(* IEC 61131-3 sources: BODAS-RC27-18_40/st/bodas_rc18_12_27_18_40/plc_logic/application/easyconfig_import/bds_out_ec, 7 files *)

(* ---- bds_out_aov_signal_te-bds_out_aov_signal_te.st ---- *)
(* --- Interface --- *)
{attribute 'qualified_only' := ''}
{attribute 'strict' := ''}
TYPE bds_out_aov_signal_te :
(
	OUT_AOV_START_SIGNALS := 16#300,
	OUT_AOV_START := 16#2FF,
	K25,
	A12,
	K62,
	OUT_AOV_NUM_SIGNALS,
	OUT_AOV_PVG_NUM_SIGNALS := K62
) UINT;
END_TYPE

(* ---- bds_out_do_signal_te-bds_out_do_signal_te.st ---- *)
(* --- Interface --- *)
{attribute 'qualified_only' := ''}
{attribute 'strict' := ''}
TYPE bds_out_do_signal_te :
(
	OUT_DO_START_SIGNALS := 16#100,
	OUT_DO_START := 16#FF,
	K13,
	A04,
	A10,
	A56,
	A11,
	A55,
	A01,
	A06,
	A16,
	A58,
	A49,
	A50,
	K84,
	K85,
	K86,
	K87,
	OUT_DO_NUM_SIGNALS,
	OUT_DO_FSC_NUM_SIGNALS := K84
) UINT;
END_TYPE

(* ---- bds_out_po_signal_te-bds_out_po_signal_te.st ---- *)
(* --- Interface --- *)
{attribute 'qualified_only' := ''}
{attribute 'strict' := ''}
TYPE bds_out_po_signal_te :
(
	OUT_PO_START_SIGNALS := 16#200,
	OUT_PO_START := 16#1FF,
	K07,
	K09,
	K73,
	K08,
	K29,
	K17,
	A32,
	A47,
	A31,
	A48,
	A46,
	A33,
	A34,
	A51,
	A35,
	A53,
	A52,
	A54,
	K16,
	K14,
	K15,
	A19,
	A05,
	A20,
	A09,
	A02,
	A17,
	K51,
	K12,
	A03,
	A18,
	A08,
	A07,
	K80,
	K81,
	K82,
	K83,
	OUT_PO_NUM_SIGNALS,
	OUT_PO_FSC_NUM_SIGNALS := K80,
	OUT_PO_FSC_HS_NUM_SIGNALS := K16
) UINT;
END_TYPE

(* ---- bds_outclcu_signal_te-bds_outClcU_signal_te.st ---- *)
(* --- Interface --- *)
{attribute 'qualified_only' := ''}
{attribute 'strict' := ''}
TYPE bds_outClcU_signal_te :
(
	bds_outClcU_K25_E := 0,
	bds_outClcU_A12_E,
	bds_outClcU_K62_E,
	bds_outClcU_numSignal_E
) USINT;
END_TYPE

(* ---- bds_outdig_signal_te-bds_outDig_signal_te.st ---- *)
(* --- Interface --- *)
{attribute 'external_name' := 'cmp_rts_bds_outDig_signal_te'}
TYPE bds_outDig_signal_te :
(
	bds_outDig_K13_E := 0,
	bds_outDig_A04_E,
	bds_outDig_A10_E,
	bds_outDig_A56_E,
	bds_outDig_A11_E,
	bds_outDig_A55_E,
	bds_outDig_A01_E,
	bds_outDig_A06_E,
	bds_outDig_A16_E,
	bds_outDig_A58_E,
	bds_outDig_A49_E,
	bds_outDig_A50_E,
	bds_outDig_K84_E,
	bds_outDig_K85_E,
	bds_outDig_K86_E,
	bds_outDig_K87_E,
	bds_outDig_K07_E,
	bds_outDig_K09_E,
	bds_outDig_K73_E,
	bds_outDig_K08_E,
	bds_outDig_K29_E,
	bds_outDig_K17_E,
	bds_outDig_A32_E,
	bds_outDig_A47_E,
	bds_outDig_A31_E,
	bds_outDig_A48_E,
	bds_outDig_A46_E,
	bds_outDig_A33_E,
	bds_outDig_A34_E,
	bds_outDig_A51_E,
	bds_outDig_A35_E,
	bds_outDig_A53_E,
	bds_outDig_A52_E,
	bds_outDig_A54_E,
	bds_outDig_K16_E,
	bds_outDig_K14_E,
	bds_outDig_K15_E,
	bds_outDig_A19_E,
	bds_outDig_A05_E,
	bds_outDig_A20_E,
	bds_outDig_A09_E,
	bds_outDig_A02_E,
	bds_outDig_A17_E,
	bds_outDig_K51_E,
	bds_outDig_K12_E,
	bds_outDig_A03_E,
	bds_outDig_A18_E,
	bds_outDig_A08_E,
	bds_outDig_A07_E,
	bds_outDig_K80_E,
	bds_outDig_K81_E,
	bds_outDig_K82_E,
	bds_outDig_K83_E,
	bds_outDig_numSignal_E
) USINT;
END_TYPE

(* ---- bds_outpwm_signal_te-bds_outPwm_signal_te.st ---- *)
(* --- Interface --- *)
{attribute 'external_name' := 'cmp_rts_bds_outPwm_signal_te'}
TYPE bds_outPwm_signal_te :
(
	bds_outPwm_K07_E := 0,
	bds_outPwm_K09_E,
	bds_outPwm_K73_E,
	bds_outPwm_K08_E,
	bds_outPwm_K29_E,
	bds_outPwm_K17_E,
	bds_outPwm_A32_E,
	bds_outPwm_A47_E,
	bds_outPwm_A31_E,
	bds_outPwm_A48_E,
	bds_outPwm_A46_E,
	bds_outPwm_A33_E,
	bds_outPwm_A34_E,
	bds_outPwm_A51_E,
	bds_outPwm_A35_E,
	bds_outPwm_A53_E,
	bds_outPwm_A52_E,
	bds_outPwm_A54_E,
	bds_outPwm_K16_E,
	bds_outPwm_K14_E,
	bds_outPwm_K15_E,
	bds_outPwm_A19_E,
	bds_outPwm_A05_E,
	bds_outPwm_A20_E,
	bds_outPwm_A09_E,
	bds_outPwm_A02_E,
	bds_outPwm_A17_E,
	bds_outPwm_K51_E,
	bds_outPwm_K12_E,
	bds_outPwm_A03_E,
	bds_outPwm_A18_E,
	bds_outPwm_A08_E,
	bds_outPwm_A07_E,
	bds_outPwm_K80_E,
	bds_outPwm_K81_E,
	bds_outPwm_K82_E,
	bds_outPwm_K83_E,
	bds_outPwm_numSignal_E
) USINT;
END_TYPE

(* ---- bds_out_ec_gvl-bds_out_ec_gvl.st ---- *)
(* --- Interface --- *)
{attribute 'qualified_only' := ''}
VAR_GLOBAL CONSTANT
	RECONF_X_X_X25: UDINT := 0;
END_VAR
